FUNCTION_BLOCK ConsoleIO (* Basic Function Block Type *)
  (* Standard: 61499-2 *)
  (* Version 0.0, 11/16/2026, Sandeep Patil, Flexbridge AB, Template *)
  PACKAGE Flexbridge.FestoMPS400;
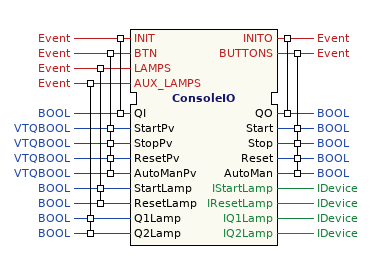
  EVENT_INPUT
    INIT WITH QI; (* Initialisation request *)
    BTN WITH StartPv, StopPv, ResetPv, AutoManPv; (* A console input changed *)
    LAMPS WITH StartLamp, ResetLamp; (* START and RESET lamps (from StationMode) *)
    AUX_LAMPS WITH Q1Lamp, Q2Lamp; (* Lamps Q1 and Q2 (from the station sequence) *)
  END_EVENT
  EVENT_OUTPUT
    INITO WITH QO; (* Initialisation confirm *)
    BUTTONS WITH Start, Stop, Reset, AutoMan; (* Button states *)
  END_EVENT
  VAR_INPUT
    QI : BOOL; (* Input event qualifier *)
    StartPv : VTQBOOL; (* S1 START button (normally open) *)
    StopPv : VTQBOOL; (* S2 STOP button (normally closed) *)
    ResetPv : VTQBOOL; (* S4 RESET button (normally open) *)
    AutoManPv : VTQBOOL; (* S3 AUTO/MAN key switch *)
    StartLamp : BOOL; (* P1 START lamp *)
    ResetLamp : BOOL; (* P2 RESET lamp *)
    Q1Lamp : BOOL; (* P3 lamp Q1 *)
    Q2Lamp : BOOL; (* P4 lamp Q2 *)
  END_VAR
  VAR_OUTPUT
    QO : BOOL; (* Output event qualifier *)
    Start : BOOL; (* START pressed *)
    Stop : BOOL; (* STOP pressed (the NC contact is inverted here) *)
    Reset : BOOL; (* RESET pressed *)
    AutoMan : BOOL; (* Key switch position *)
  END_VAR
  PLUGS
    IStartLamp : IDevice;
    IResetLamp : IDevice;
    IQ1Lamp : IDevice;
    IQ2Lamp : IDevice;
  END_PLUGS
  VAR
    CurStartLamp : BOOL; (* StartLamp as last commanded *)
    CurResetLamp : BOOL; (* ResetLamp as last commanded *)
    CurQ1Lamp : BOOL; (* Q1Lamp as last commanded *)
    CurQ2Lamp : BOOL; (* Q2Lamp as last commanded *)
    ChStartLamp : BOOL; (* StartLamp changed at this event *)
    ChResetLamp : BOOL; (* ResetLamp changed at this event *)
    ChQ1Lamp : BOOL; (* Q1Lamp changed at this event *)
    ChQ2Lamp : BOOL; (* Q2Lamp changed at this event *)
    ReqStartLamp : BOOL; (* StartLamp as requested before INIT *)
    ReqResetLamp : BOOL; (* ResetLamp as requested before INIT *)
    ReqQ1Lamp : BOOL; (* Q1Lamp as requested before INIT *)
    ReqQ2Lamp : BOOL; (* Q2Lamp as requested before INIT *)
    SyncedStartLamp : BOOL; (* StartLamp has received its state while program local *)
    SyncedResetLamp : BOOL; (* ResetLamp has received its state while program local *)
    SyncedQ1Lamp : BOOL; (* Q1Lamp has received its state while program local *)
    SyncedQ2Lamp : BOOL; (* Q2Lamp has received its state while program local *)
    TriesStartLamp : INT; (* Program-local requests sent to StartLamp after a ready report *)
    TriesResetLamp : INT; (* Program-local requests sent to ResetLamp after a ready report *)
    TriesQ1Lamp : INT; (* Program-local requests sent to Q1Lamp after a ready report *)
    TriesQ2Lamp : INT; (* Program-local requests sent to Q2Lamp after a ready report *)
    NeedSel : BOOL; (* The lamp that just reported ready must be switched to program local *)
  END_VAR
  EC_STATES
    START; (* Initial state: not initialised yet, lamp requests are stored *)
    PRE_LMP : algStoreLamps;
    PRE_AUX : algStoreAux;
    INIT_S : algInit, -> IStartLamp.REQ_CMD, -> IResetLamp.REQ_CMD, -> IQ1Lamp.REQ_CMD, -> IQ2Lamp.REQ_CMD, -> INITO;
    READY; (* Initialised *)
    BTN_S : algButtons -> BUTTONS;
    LMP_S : algLamps;
    LMP_START : -> IStartLamp.REQ_CMD;
    LMP_C2;
    LMP_RESET : -> IResetLamp.REQ_CMD;
    AUX_S : algAuxLamps;
    AUX_Q1 : -> IQ1Lamp.REQ_CMD;
    AUX_C2;
    AUX_Q2 : -> IQ2Lamp.REQ_CMD;
    RDY_StartLamp : algReadyStartLamp;
    SEL_StartLamp : -> IStartLamp.REQ_PROGLOCALSEL, -> IStartLamp.REQ_CMD;
    RDY_ResetLamp : algReadyResetLamp;
    SEL_ResetLamp : -> IResetLamp.REQ_PROGLOCALSEL, -> IResetLamp.REQ_CMD;
    RDY_Q1Lamp : algReadyQ1Lamp;
    SEL_Q1Lamp : -> IQ1Lamp.REQ_PROGLOCALSEL, -> IQ1Lamp.REQ_CMD;
    RDY_Q2Lamp : algReadyQ2Lamp;
    SEL_Q2Lamp : -> IQ2Lamp.REQ_PROGLOCALSEL, -> IQ2Lamp.REQ_CMD;
  END_STATES
  EC_TRANSITIONS
    START TO INIT_S := INIT;
    START TO PRE_LMP := LAMPS;
    PRE_LMP TO START := 1;
    START TO PRE_AUX := AUX_LAMPS;
    PRE_AUX TO START := 1;
    INIT_S TO READY := 1;
    READY TO INIT_S := INIT;
    READY TO BTN_S := BTN;
    BTN_S TO READY := 1;
    READY TO LMP_S := LAMPS;
    LMP_S TO LMP_START := ChStartLamp;
    LMP_S TO LMP_C2 := NOT ChStartLamp;
    LMP_START TO LMP_C2 := 1;
    LMP_C2 TO LMP_RESET := ChResetLamp;
    LMP_C2 TO READY := NOT ChResetLamp;
    LMP_RESET TO READY := 1;
    READY TO AUX_S := AUX_LAMPS;
    AUX_S TO AUX_Q1 := ChQ1Lamp;
    AUX_S TO AUX_C2 := NOT ChQ1Lamp;
    AUX_Q1 TO AUX_C2 := 1;
    AUX_C2 TO AUX_Q2 := ChQ2Lamp;
    AUX_C2 TO READY := NOT ChQ2Lamp;
    AUX_Q2 TO READY := 1;
    READY TO RDY_StartLamp := IStartLamp.CNF_READY;
    RDY_StartLamp TO SEL_StartLamp := NeedSel;
    RDY_StartLamp TO READY := NOT NeedSel;
    SEL_StartLamp TO READY := 1;
    READY TO RDY_ResetLamp := IResetLamp.CNF_READY;
    RDY_ResetLamp TO SEL_ResetLamp := NeedSel;
    RDY_ResetLamp TO READY := NOT NeedSel;
    SEL_ResetLamp TO READY := 1;
    READY TO RDY_Q1Lamp := IQ1Lamp.CNF_READY;
    RDY_Q1Lamp TO SEL_Q1Lamp := NeedSel;
    RDY_Q1Lamp TO READY := NOT NeedSel;
    SEL_Q1Lamp TO READY := 1;
    READY TO RDY_Q2Lamp := IQ2Lamp.CNF_READY;
    RDY_Q2Lamp TO SEL_Q2Lamp := NeedSel;
    RDY_Q2Lamp TO READY := NOT NeedSel;
    SEL_Q2Lamp TO READY := 1;
  END_TRANSITIONS
  ALGORITHM algInit IN ST: (* Apply the lamp states requested so far (program local is selected on CNF_READY) *)
QO := QI;
IStartLamp.ProgLocalSel := TRUE;
IF ReqStartLamp THEN IStartLamp.Lsp.value := 1; ELSE IStartLamp.Lsp.value := 0; END_IF;
CurStartLamp := ReqStartLamp;
IResetLamp.ProgLocalSel := TRUE;
IF ReqResetLamp THEN IResetLamp.Lsp.value := 1; ELSE IResetLamp.Lsp.value := 0; END_IF;
CurResetLamp := ReqResetLamp;
IQ1Lamp.ProgLocalSel := TRUE;
IF ReqQ1Lamp THEN IQ1Lamp.Lsp.value := 1; ELSE IQ1Lamp.Lsp.value := 0; END_IF;
CurQ1Lamp := ReqQ1Lamp;
IQ2Lamp.ProgLocalSel := TRUE;
IF ReqQ2Lamp THEN IQ2Lamp.Lsp.value := 1; ELSE IQ2Lamp.Lsp.value := 0; END_IF;
CurQ2Lamp := ReqQ2Lamp;
  END_ALGORITHM
  ALGORITHM algStoreLamps IN ST: (* Before INIT: remember the START and RESET lamp request *)
ReqStartLamp := StartLamp;
ReqResetLamp := ResetLamp;
  END_ALGORITHM
  ALGORITHM algStoreAux IN ST: (* Before INIT: remember the Q1 and Q2 lamp request *)
ReqQ1Lamp := Q1Lamp;
ReqQ2Lamp := Q2Lamp;
  END_ALGORITHM
  ALGORITHM algButtons IN ST: (* Button states from the inputs; STOP is a normally closed contact *)
Start := StartPv.value;
Stop := NOT StopPv.value;
Reset := ResetPv.value;
AutoMan := AutoManPv.value;
  END_ALGORITHM
  ALGORITHM algLamps IN ST: (* START and RESET lamps: command only those that changed *)
ChStartLamp := StartLamp <> CurStartLamp;
CurStartLamp := StartLamp;
IF StartLamp THEN IStartLamp.Lsp.value := 1; ELSE IStartLamp.Lsp.value := 0; END_IF;
ChResetLamp := ResetLamp <> CurResetLamp;
CurResetLamp := ResetLamp;
IF ResetLamp THEN IResetLamp.Lsp.value := 1; ELSE IResetLamp.Lsp.value := 0; END_IF;
  END_ALGORITHM
  ALGORITHM algAuxLamps IN ST: (* Lamps Q1 and Q2: command only those that changed *)
ChQ1Lamp := Q1Lamp <> CurQ1Lamp;
CurQ1Lamp := Q1Lamp;
IF Q1Lamp THEN IQ1Lamp.Lsp.value := 1; ELSE IQ1Lamp.Lsp.value := 0; END_IF;
ChQ2Lamp := Q2Lamp <> CurQ2Lamp;
CurQ2Lamp := Q2Lamp;
IF Q2Lamp THEN IQ2Lamp.Lsp.value := 1; ELSE IQ2Lamp.Lsp.value := 0; END_IF;
  END_ALGORITHM
  ALGORITHM algReadyStartLamp IN ST: (* StartLamp reported ready: send owner request and lamp state again until synchronised *)
NeedSel := NOT SyncedStartLamp AND TriesStartLamp < 3;
IF NeedSel THEN
    TriesStartLamp := TriesStartLamp + 1;
    IStartLamp.ProgLocalSel := TRUE;
    IF CurStartLamp THEN IStartLamp.Lsp.value := 1; ELSE IStartLamp.Lsp.value := 0; END_IF;
    SyncedStartLamp := IStartLamp.ProgLocal;
END_IF;
  END_ALGORITHM
  ALGORITHM algReadyResetLamp IN ST: (* ResetLamp reported ready: send owner request and lamp state again until synchronised *)
NeedSel := NOT SyncedResetLamp AND TriesResetLamp < 3;
IF NeedSel THEN
    TriesResetLamp := TriesResetLamp + 1;
    IResetLamp.ProgLocalSel := TRUE;
    IF CurResetLamp THEN IResetLamp.Lsp.value := 1; ELSE IResetLamp.Lsp.value := 0; END_IF;
    SyncedResetLamp := IResetLamp.ProgLocal;
END_IF;
  END_ALGORITHM
  ALGORITHM algReadyQ1Lamp IN ST: (* Q1Lamp reported ready: send owner request and lamp state again until synchronised *)
NeedSel := NOT SyncedQ1Lamp AND TriesQ1Lamp < 3;
IF NeedSel THEN
    TriesQ1Lamp := TriesQ1Lamp + 1;
    IQ1Lamp.ProgLocalSel := TRUE;
    IF CurQ1Lamp THEN IQ1Lamp.Lsp.value := 1; ELSE IQ1Lamp.Lsp.value := 0; END_IF;
    SyncedQ1Lamp := IQ1Lamp.ProgLocal;
END_IF;
  END_ALGORITHM
  ALGORITHM algReadyQ2Lamp IN ST: (* Q2Lamp reported ready: send owner request and lamp state again until synchronised *)
NeedSel := NOT SyncedQ2Lamp AND TriesQ2Lamp < 3;
IF NeedSel THEN
    TriesQ2Lamp := TriesQ2Lamp + 1;
    IQ2Lamp.ProgLocalSel := TRUE;
    IF CurQ2Lamp THEN IQ2Lamp.Lsp.value := 1; ELSE IQ2Lamp.Lsp.value := 0; END_IF;
    SyncedQ2Lamp := IQ2Lamp.ProgLocal;
END_IF;
  END_ALGORITHM
END_FUNCTION_BLOCK
